// TIA Portal V21 export
// export: Created 2026-11-22T02:34:37.0667875Z, ExportSetting WithDefaults, DisplayName Totally Integrated Automation Portal, DisplayVersion V21 Update 3, DisplayName STEP 7 Professional, DisplayVersion V21 Update 3, DisplayName STEP 7 Safety, DisplayVersion V21, DisplayName Tech WebApplication, DisplayVersion V21, DisplayName WinCC Basic/Comfort/Advanced, DisplayVersion V21 Update 3, DisplayName WinCC Unified, DisplayVersion V21 Update 3
VBScript "SetS4"  Type=Sub
  SmartTags("D_State") = 4
  SmartTags("D_Bool") = False
  SmartTags("D_SInt") = -1
  SmartTags("D_Int") = -1
  SmartTags("D_DInt") = 0
  SmartTags("D_USInt") = 1
  SmartTags("D_UInt") = 1
  SmartTags("D_UDInt") = 1
  SmartTags("D_Real") = 0.0005
  SmartTags("D_LReal") = -0.0
  SmartTags("D_String") = "äöü ÄÖÜ ß"
  SmartTags("D_DateTime") = DateSerial(1970, 1, 1) + TimeSerial(0, 0, 0)
  SmartTags("D_Pct") = 150
  SmartTags("D_Range") = 200
  SmartTags("D_Bits") = 9
  SmartTags("D_Vis") = False
  SmartTags("D_En") = True
  SmartTags("D_X") = -20
  SmartTags("D_Y") = 0
  SmartTags("D_Max") = 100
  SmartTags("D_Min") = 0
  SmartTags("D_TL") = 50
  SmartTags("D_BarR") = 2.5
